// TIA Portal V21 export
// export: Created 2026-11-10T07:27:31.0404088Z, ExportSetting WithDefaults, DisplayName Totally Integrated Automation Portal, DisplayVersion V21 Update 3, DisplayName STEP 7 Professional, DisplayVersion V21 Update 3, DisplayName STEP 7 Safety, DisplayVersion V21, DisplayName Tech WebApplication, DisplayVersion V21, DisplayName WinCC Basic/Comfort/Advanced, DisplayVersion V21 Update 3, DisplayName WinCC Unified, DisplayVersion V21 Update 3
FUNCTION_BLOCK "FB_SclTech"   // FB7, SCL
{ S7_Optimized_Access := 'TRUE' }
VERSION : 0.1
// stored: AutoNumber true, IsIECCheckEnabled false, IsRetainMemResEnabled false, MemoryReserve 100, SetENOAutomatically false, UDAEnableTagReadback false
   VAR_INPUT
      sp : Real;
      pv : Real;
   END_VAR
   VAR_OUTPUT
      outv : Real;
      err : Bool;
   END_VAR
BEGIN
// PID call
   "PID_Comp_2_3"(Setpoint := #sp, Input := #pv, Output => #outv, Error => #err);
END_FUNCTION_BLOCK
